% RSLogix 500 project PROYECTO1_TEST.RSS, saved by version 12.00.00.00 %
PROJECT "UNTITLED"    % processor: SLC 500, 1747-L541 %

PROGRAM FILES
  LAD 2   26 rungs

DATA FILES
  O0   33 elements
  I1   33 elements
  S2   164 elements
  B3   4 elements
  T4   6 elements
  C5   1 elements
  R6   1 elements
  N7   4 elements
  F8   1 elements

LADDER 2
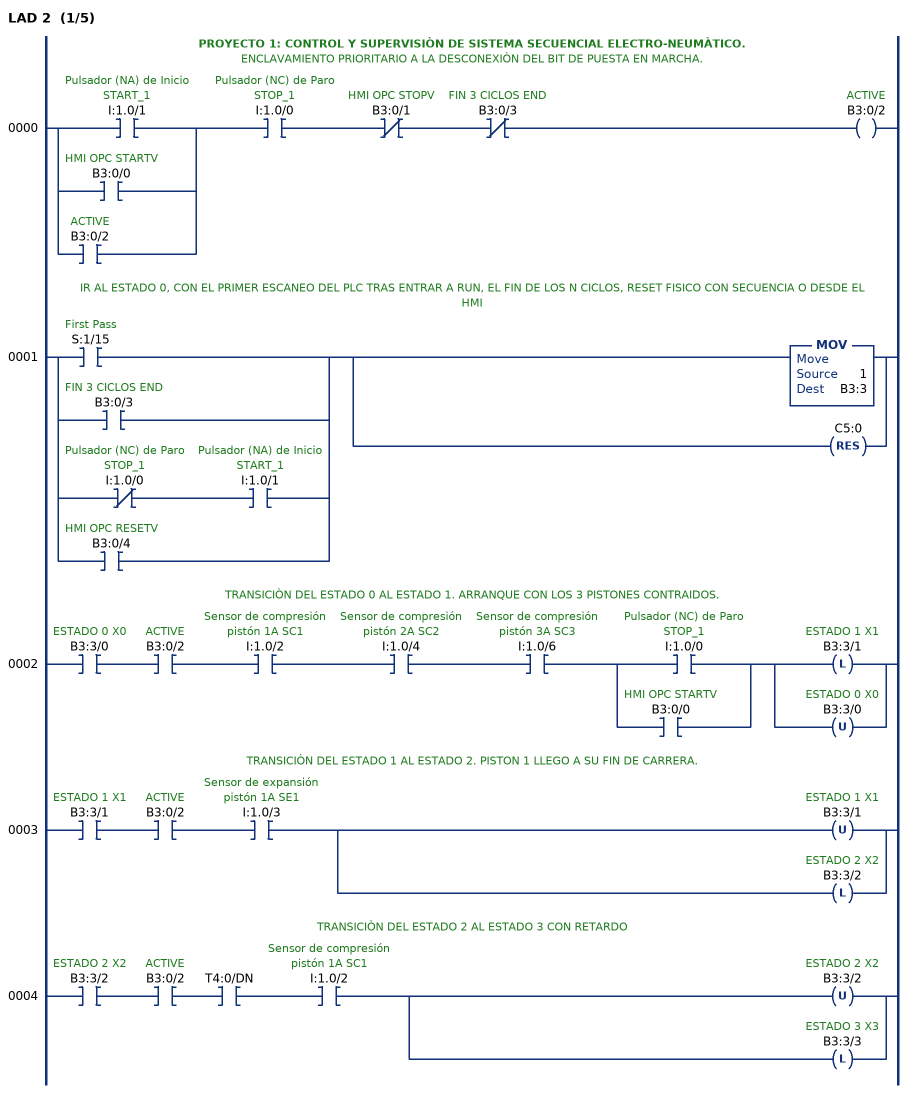
% Rung: 0 %
% TITLE: PROYECTO 1: CONTROL Y SUPERVISIÒN DE SISTEMA SECUENCIAL ELECTRO-NEUMÀTICO. %
% ENCLAVAMIENTO PRIORITARIO A LA DESCONEXIÒN DEL BIT DE PUESTA EN MARCHA. %
SOR BST XIC I:1.0/1 NXB XIC B3:0/0 NXB XIC B3:0/2 BND XIC I:1.0/0 XIO B3:0/1 XIO B3:0/3 OTE B3:0/2 EOR
%   I:1.0/1  START_1  "Pulsador (NA) de Inicio" %
%   B3:0/0  STARTV  "HMI OPC" %
%   B3:0/2  ACTIVE %
%   I:1.0/0  STOP_1  "Pulsador (NC) de Paro" %
%   B3:0/1  STOPV  "HMI OPC" %
%   B3:0/3  END  "FIN 3 CICLOS" %
% Rung: 1 %
% IR AL ESTADO 0, CON EL PRIMER ESCANEO DEL PLC TRAS ENTRAR A RUN, EL FIN DE LOS N CICLOS, RESET FISICO CON SECUENCIA O DESDE EL HMI %
SOR BST XIC S:1/15 NXB XIC B3:0/3 NXB XIO I:1.0/0 XIC I:1.0/1 NXB XIC B3:0/4 BND BST MOV 1 B3:3 NXB RES C5:0 BND EOR
%   S:1/15  "First Pass" %
%   B3:0/3  END  "FIN 3 CICLOS" %
%   I:1.0/0  STOP_1  "Pulsador (NC) de Paro" %
%   I:1.0/1  START_1  "Pulsador (NA) de Inicio" %
%   B3:0/4  RESETV  "HMI OPC" %
% Rung: 2 %
% TRANSICIÒN DEL ESTADO 0 AL ESTADO 1. ARRANQUE CON LOS 3 PISTONES CONTRAIDOS. %
SOR XIC B3:3/0 XIC B3:0/2 XIC I:1.0/2 XIC I:1.0/4 XIC I:1.0/6 BST XIC I:1.0/0 NXB XIC B3:0/0 BND BST OTL B3:3/1 NXB OTU B3:3/0 BND EOR
%   B3:3/0  X0  "ESTADO 0" %
%   B3:0/2  ACTIVE %
%   I:1.0/2  SC1  "Sensor de compresión pistón 1A" %
%   I:1.0/4  SC2  "Sensor de compresión pistón 2A" %
%   I:1.0/6  SC3  "Sensor de compresión pistón 3A" %
%   I:1.0/0  STOP_1  "Pulsador (NC) de Paro" %
%   B3:0/0  STARTV  "HMI OPC" %
%   B3:3/1  X1  "ESTADO 1" %
% Rung: 3 %
% TRANSICIÒN DEL ESTADO 1 AL ESTADO 2. PISTON 1 LLEGO A SU FIN DE CARRERA. %
SOR XIC B3:3/1 XIC B3:0/2 XIC I:1.0/3 BST OTU B3:3/1 NXB OTL B3:3/2 BND EOR
%   B3:3/1  X1  "ESTADO 1" %
%   B3:0/2  ACTIVE %
%   I:1.0/3  SE1  "Sensor de expansión pistón 1A" %
%   B3:3/2  X2  "ESTADO 2" %
% Rung: 4 %
% TRANSICIÒN DEL ESTADO 2 AL ESTADO 3 CON RETARDO %
SOR XIC B3:3/2 XIC B3:0/2 XIC T4:0/DN XIC I:1.0/2 BST OTU B3:3/2 NXB OTL B3:3/3 BND EOR
%   B3:3/2  X2  "ESTADO 2" %
%   B3:0/2  ACTIVE %
%   I:1.0/2  SC1  "Sensor de compresión pistón 1A" %
%   B3:3/3  X3  "ESTADO 3" %

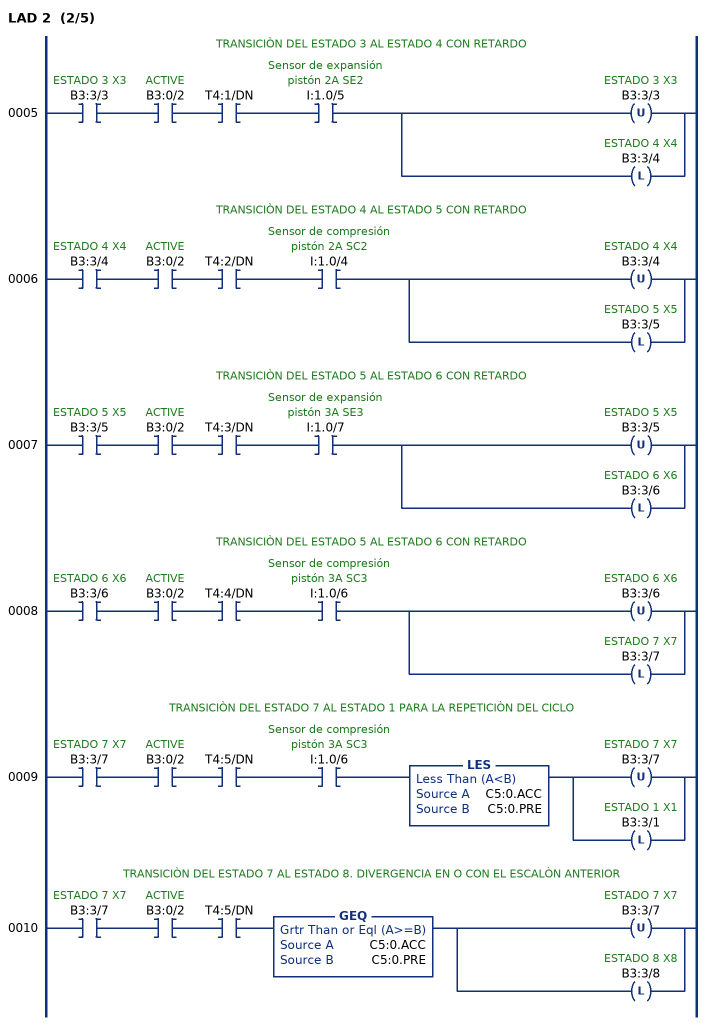
% Rung: 5 %
% TRANSICIÒN DEL ESTADO 3 AL ESTADO 4 CON RETARDO %
SOR XIC B3:3/3 XIC B3:0/2 XIC T4:1/DN XIC I:1.0/5 BST OTU B3:3/3 NXB OTL B3:3/4 BND EOR
%   B3:3/3  X3  "ESTADO 3" %
%   B3:0/2  ACTIVE %
%   I:1.0/5  SE2  "Sensor de expansión pistón 2A" %
%   B3:3/4  X4  "ESTADO 4" %
% Rung: 6 %
% TRANSICIÒN DEL ESTADO 4 AL ESTADO 5 CON RETARDO %
SOR XIC B3:3/4 XIC B3:0/2 XIC T4:2/DN XIC I:1.0/4 BST OTU B3:3/4 NXB OTL B3:3/5 BND EOR
%   B3:3/4  X4  "ESTADO 4" %
%   B3:0/2  ACTIVE %
%   I:1.0/4  SC2  "Sensor de compresión pistón 2A" %
%   B3:3/5  X5  "ESTADO 5" %
% Rung: 7 %
% TRANSICIÒN DEL ESTADO 5 AL ESTADO 6 CON RETARDO %
SOR XIC B3:3/5 XIC B3:0/2 XIC T4:3/DN XIC I:1.0/7 BST OTU B3:3/5 NXB OTL B3:3/6 BND EOR
%   B3:3/5  X5  "ESTADO 5" %
%   B3:0/2  ACTIVE %
%   I:1.0/7  SE3  "Sensor de expansión pistón 3A" %
%   B3:3/6  X6  "ESTADO 6" %
% Rung: 8 %
% TRANSICIÒN DEL ESTADO 5 AL ESTADO 6 CON RETARDO %
SOR XIC B3:3/6 XIC B3:0/2 XIC T4:4/DN XIC I:1.0/6 BST OTU B3:3/6 NXB OTL B3:3/7 BND EOR
%   B3:3/6  X6  "ESTADO 6" %
%   B3:0/2  ACTIVE %
%   I:1.0/6  SC3  "Sensor de compresión pistón 3A" %
%   B3:3/7  X7  "ESTADO 7" %
% Rung: 9 %
% TRANSICIÒN DEL ESTADO 7 AL ESTADO 1 PARA LA REPETICIÒN DEL CICLO %
SOR XIC B3:3/7 XIC B3:0/2 XIC T4:5/DN XIC I:1.0/6 LES C5:0.ACC C5:0.PRE BST OTU B3:3/7 NXB OTL B3:3/1 BND EOR
%   B3:3/7  X7  "ESTADO 7" %
%   B3:0/2  ACTIVE %
%   I:1.0/6  SC3  "Sensor de compresión pistón 3A" %
%   B3:3/1  X1  "ESTADO 1" %
% Rung: 10 %
% TRANSICIÒN DEL ESTADO 7 AL ESTADO 8. DIVERGENCIA EN O CON EL ESCALÒN ANTERIOR %
SOR XIC B3:3/7 XIC B3:0/2 XIC T4:5/DN GEQ C5:0.ACC C5:0.PRE BST OTU B3:3/7 NXB OTL B3:3/8 BND EOR
%   B3:3/7  X7  "ESTADO 7" %
%   B3:0/2  ACTIVE %
%   B3:3/8  X8  "ESTADO 8" %

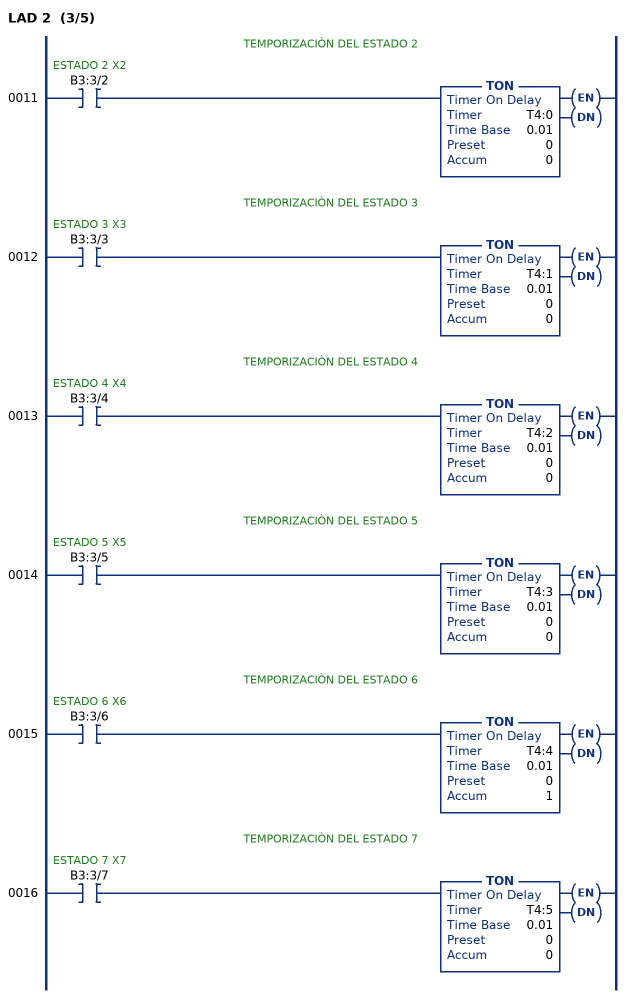
% Rung: 11 %
% TEMPORIZACIÒN DEL ESTADO 2 %
SOR XIC B3:3/2 TON T4:0 0.01 0 0 EOR
%   B3:3/2  X2  "ESTADO 2" %
% Rung: 12 %
% TEMPORIZACIÒN DEL ESTADO 3 %
SOR XIC B3:3/3 TON T4:1 0.01 0 0 EOR
%   B3:3/3  X3  "ESTADO 3" %
% Rung: 13 %
% TEMPORIZACIÒN DEL ESTADO 4 %
SOR XIC B3:3/4 TON T4:2 0.01 0 0 EOR
%   B3:3/4  X4  "ESTADO 4" %
% Rung: 14 %
% TEMPORIZACIÒN DEL ESTADO 5 %
SOR XIC B3:3/5 TON T4:3 0.01 0 0 EOR
%   B3:3/5  X5  "ESTADO 5" %
% Rung: 15 %
% TEMPORIZACIÒN DEL ESTADO 6 %
SOR XIC B3:3/6 TON T4:4 0.01 0 1 EOR
%   B3:3/6  X6  "ESTADO 6" %
% Rung: 16 %
% TEMPORIZACIÒN DEL ESTADO 7 %
SOR XIC B3:3/7 TON T4:5 0.01 0 0 EOR
%   B3:3/7  X7  "ESTADO 7" %

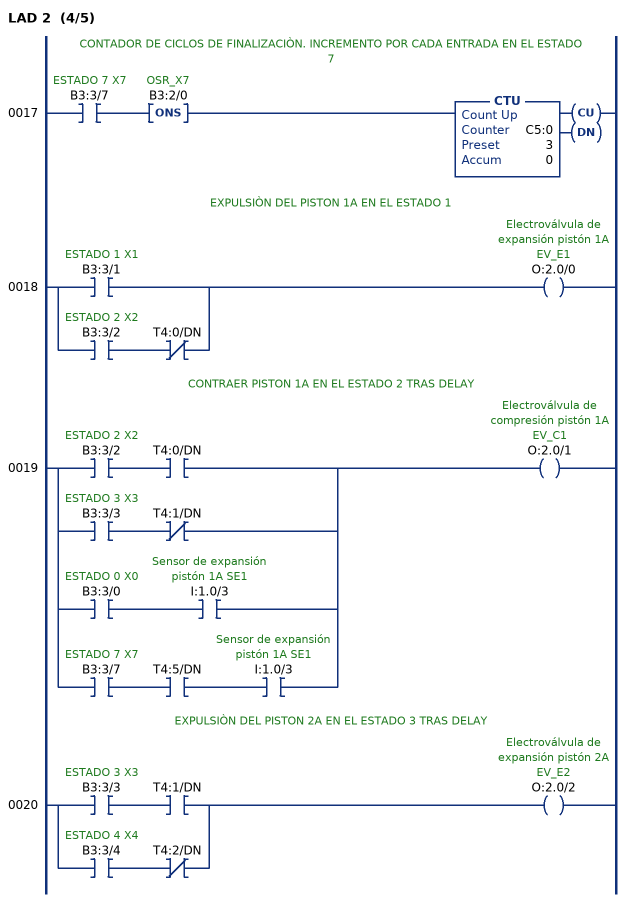
% Rung: 17 %
% CONTADOR DE CICLOS DE FINALIZACIÒN. INCREMENTO POR CADA ENTRADA EN EL ESTADO 7 %
SOR XIC B3:3/7 OSR B3:2/0 CTU C5:0 3 0 EOR
%   B3:3/7  X7  "ESTADO 7" %
%   B3:2/0  OSR_X7 %
% Rung: 18 %
% EXPULSIÒN DEL PISTON 1A EN EL ESTADO 1 %
SOR BST XIC B3:3/1 NXB XIC B3:3/2 XIO T4:0/DN BND OTE O:2.0/0 EOR
%   B3:3/1  X1  "ESTADO 1" %
%   B3:3/2  X2  "ESTADO 2" %
%   O:2.0/0  EV_E1  "Electroválvula de expansión pistón 1A" %
% Rung: 19 %
% CONTRAER PISTON 1A EN EL ESTADO 2 TRAS DELAY %
SOR BST XIC B3:3/2 XIC T4:0/DN NXB XIC B3:3/3 XIO T4:1/DN NXB XIC B3:3/0 XIC I:1.0/3 NXB XIC B3:3/7 XIC T4:5/DN XIC I:1.0/3 BND OTE O:2.0/1 EOR
%   B3:3/2  X2  "ESTADO 2" %
%   B3:3/3  X3  "ESTADO 3" %
%   B3:3/0  X0  "ESTADO 0" %
%   I:1.0/3  SE1  "Sensor de expansión pistón 1A" %
%   B3:3/7  X7  "ESTADO 7" %
%   O:2.0/1  EV_C1  "Electroválvula de compresión pistón 1A" %
% Rung: 20 %
% EXPULSIÒN DEL PISTON 2A EN EL ESTADO 3 TRAS DELAY %
SOR BST XIC B3:3/3 XIC T4:1/DN NXB XIC B3:3/4 XIO T4:2/DN BND OTE O:2.0/2 EOR
%   B3:3/3  X3  "ESTADO 3" %
%   B3:3/4  X4  "ESTADO 4" %
%   O:2.0/2  EV_E2  "Electroválvula de expansión pistón 2A" %

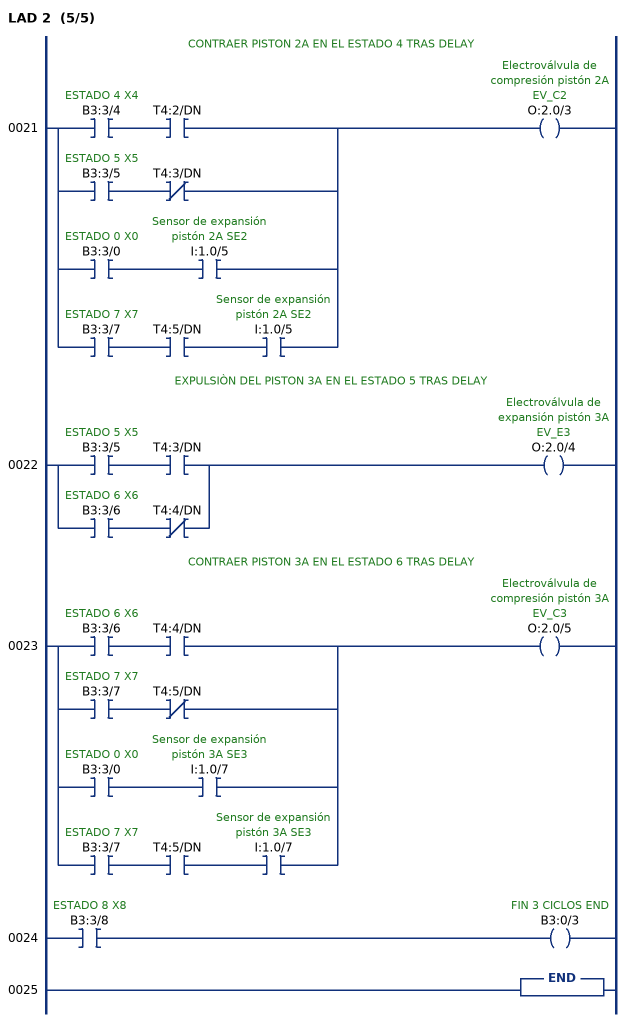
% Rung: 21 %
% CONTRAER PISTON 2A EN EL ESTADO 4 TRAS DELAY %
SOR BST XIC B3:3/4 XIC T4:2/DN NXB XIC B3:3/5 XIO T4:3/DN NXB XIC B3:3/0 XIC I:1.0/5 NXB XIC B3:3/7 XIC T4:5/DN XIC I:1.0/5 BND OTE O:2.0/3 EOR
%   B3:3/4  X4  "ESTADO 4" %
%   B3:3/5  X5  "ESTADO 5" %
%   B3:3/0  X0  "ESTADO 0" %
%   I:1.0/5  SE2  "Sensor de expansión pistón 2A" %
%   B3:3/7  X7  "ESTADO 7" %
%   O:2.0/3  EV_C2  "Electroválvula de compresión pistón 2A" %
% Rung: 22 %
% EXPULSIÒN DEL PISTON 3A EN EL ESTADO 5 TRAS DELAY %
SOR BST XIC B3:3/5 XIC T4:3/DN NXB XIC B3:3/6 XIO T4:4/DN BND OTE O:2.0/4 EOR
%   B3:3/5  X5  "ESTADO 5" %
%   B3:3/6  X6  "ESTADO 6" %
%   O:2.0/4  EV_E3  "Electroválvula de expansión pistón 3A" %
% Rung: 23 %
% CONTRAER PISTON 3A EN EL ESTADO 6 TRAS DELAY %
SOR BST XIC B3:3/6 XIC T4:4/DN NXB XIC B3:3/7 XIO T4:5/DN NXB XIC B3:3/0 XIC I:1.0/7 NXB XIC B3:3/7 XIC T4:5/DN XIC I:1.0/7 BND OTE O:2.0/5 EOR
%   B3:3/6  X6  "ESTADO 6" %
%   B3:3/7  X7  "ESTADO 7" %
%   B3:3/0  X0  "ESTADO 0" %
%   I:1.0/7  SE3  "Sensor de expansión pistón 3A" %
%   O:2.0/5  EV_C3  "Electroválvula de compresión pistón 3A" %
% Rung: 24 %
SOR XIC B3:3/8 OTE B3:0/3 EOR
%   B3:3/8  X8  "ESTADO 8" %
%   B3:0/3  END  "FIN 3 CICLOS" %
% Rung: 25 %
SOR END EOR

OTHER DOCUMENTED ADDRESSES
  C5:0/CU  C_CICLOS  "CICLOS"
  O:3.0/1  EV_C11  "SOLENOIDE 1A-"
  O:3.0/2  EV_E21  "SOLENOIDE 2A+"
  O:3.0/3  EV_C21  "SOLENOIDE 2A-"
  O:3.0/4  EV_E31  "SOLENOIDE 3A+"
  O:3.0/5  EV_C31  "SOLENOIDE 3A-"

COMMENTS NOT ATTACHED TO A CURRENT RUNG
  O:2.0/0: PROYECTO 1: CONTROL Y SUPERVISIÒN DE SISTEMA SECUENCIAL ELECTRO-NEUMÀTICO. / ENCLAVAMIENTO PRIORITARIO A LA DESCONEXIÒN DEL BIT DE PUESTA EN MARCHA.

DATA TABLE (non-zero values as saved)
DATA B3
% B3:0 % 0X0000 0X0000 0X0000 0X0040
DATA T4
% .PRE .ACC %
% T4:4 % 0 1
DATA C5
% .PRE .ACC %
% C5:0 % 3 0
DATA N7
% N7:0 % 0 3 0 0
